Staubli VAL3: IHM.pgx

program IHM()
begin
  userPage("IHM")
  while true
    delay(0.5)
  endWhile
end
